(* IEC 61131-3 sources: codesys-framework/txt/application/WeVe Core (library)/10 Mode/DUT, 2 files *)

(* ---- E_DefaultModes.dut.st ---- *)
{attribute 'qualified_only'}
{attribute 'strict'}
TYPE E_DefaultModes :
(
	Auto := 0,
	Manual,
	Maintenance,
	UserDefined1,
	UserDefined2,
	UserDefined3,
	UserDefined4,
	UserDefined5,
	UserDefined6,
	UserDefined7,
	UserDefined8,
	UserDefined9,
	UserDefined10
)USINT;
END_TYPE

(* ---- E_ModeStates.dut.st ---- *)
{attribute 'qualified_only'}
{attribute 'strict'}
TYPE E_ModeStates :
(
	Off := 0,
	Invalid,
	Initialize,
	Standby,
	Starting,
	Run,
	Stop,
	QuickStop,
	Safe,
	Reset
)USINT;
END_TYPE
